Fanuc KAREL source: kb00086.KL

-- PROVISIONAL review KL for V940-1; original PC SHA256 23ac743ef25d3b16abea1264f99e444cb46e8e5da154269d143c3f5861a7df84
-- Incomplete behavior may be omitted. Consult companion uncertainty JSON. Do not deploy.
PROGRAM KB00086
%NOLOCKGROUP
BEGIN
  -- V9_ZERO_TABLE_METADATA_HINT layout=0002_ascii; no indexed target words; source/name/runtime held
  -- UNRESOLVED_PC offsets 5-12; opcodes 9D,23
  -- UNRESOLVED_PC offsets 17-24; opcodes 9D,23
  -- UNRESOLVED_PC offsets 29-36; opcodes 9D,23
  -- UNRESOLVED_PC offsets 41-48; opcodes 9D,23
  -- UNRESOLVED_PC offsets 53-60; opcodes 9D,23
  -- UNRESOLVED_PC offsets 65-72; opcodes 9D,23
  -- UNRESOLVED_PC offsets 77-117; opcodes 27,22,22,22,22,22,22,31
  -- UNRESOLVED_PC offsets 122-126; opcodes 7F
END KB00086
